FUNCTION_BLOCK FB_FuseControl
VAR_INPUT
	bResetChannels:	BOOL;
END_VAR
VAR_OUTPUT
	fbError:		FB_Error;
END_VAR
VAR
	fbBlockFuse:	FB_BlockEconomySmart;
	nChannel:		INT;
END_VAR

fbBlockFuse();
FOR nChannel := fbBlockFuse.MIN_CHANNEL TO fbBlockFuse.MAX_CHANNEL DO
	CASE fbBlockFuse.Status[nChannel] OF 
		fbBlockFuse.STATUS_TRIP:
			fbError.M_Set(1, CONCAT('Sicherung hat ausgelöst! Kanal ', TO_STRING(nChannel)), 0, E_ErrorIDs.eFuseTripped, E_ErrorSrcs.eFuse);
			EXIT;
		fbBlockFuse.STATUS_OVERCURRENT:
			fbError.M_Set(1, CONCAT('Sicherung Überstrom! Kanal ', TO_STRING(nChannel)), 0, E_ErrorIDs.eFuseOvercurrent, E_ErrorSrcs.eFuse);
			EXIT;
		fbBlockFuse.STATUS_OFF:
			fbError.M_Set(1, CONCAT('Sicherung ausgeschaltet! Kanal ', TO_STRING(nChannel)), 0, E_ErrorIDs.eFuseOff, E_ErrorSrcs.eFuse);
			EXIT;
		fbBlockFuse.STATUS_ON:
			IF fbError.bError THEN
				fbError.M_Reset();				
			END_IF
		ELSE
			fbError.M_Set(1, CONCAT('Sicherung ausgeschaltet! Kanal ', TO_STRING(nChannel)), 0, E_ErrorIDs.eFuseOff, E_ErrorSrcs.eFuse);
			EXIT;
	END_CASE
END_FOR

IF fbBlockFuse.FuseTripped AND bResetChannels THEN
	fbBlockFuse.reset();
END_IF

END_FUNCTION_BLOCK

(* stored: Version 1.1.0.1, ProductVersion 3.1.4024.12
   POU FB_FuseControl: Id {5274ca77-2d19-495b-afdf-f0f4c9c09e36}, SpecialFunc None *)
